GLOBALCONSTANTS OpcUaLokal (* OPC-UA-IDs fuer die lokalen Uebungen (ein Geraet) *)
  (* Standard: 61499-1; Description: Copyright (c) 2026 Meisterschulen am Ostbahnhof This program and the accompanying materials are made available under the terms of the Eclipse Public License 2.0 which is available at https://www.eclipse.org/legal/epl-2.0/ SPDX-License-Identifier: EPL-2.0 *)
  (* Version 1.0, 2026-10-18, Franz Höpfinger, Meisterschulen am Ostbahnhof, Lokal: READ/WRITE/CREATE_METHOD ohne Endpunkt, CALL_METHOD per localhost *)
  PACKAGE Meins::OPC_UA_Lokal::const;
  VAR_GLOBAL CONSTANT
    LOCAL_OPC : WSTRING := "opc.tcp://localhost:4840"; (* Eigener Server (localhost), nur fuer CALL_METHOD *)
    L01_Q1_NODE : WSTRING := "/Objects/Lokal/L01/Q1,1:s=L01_Q1"; (* L01: Knoten Q1 *)
    L01_Q1_WRITE : WSTRING := MyLib_OPC::F_OPC_LOCAL("WRITE", L01_Q1_NODE); (* L01: Input_I1 schreibt lokal (PUBLISH) *)
    L01_Q1_READ : WSTRING := MyLib_OPC::F_OPC_LOCAL("READ", L01_Q1_NODE); (* L01: Output_Q1 liest lokal (SUBSCRIBE) *)
    L03_FF1_TRIGGER_NODE : WSTRING := "/Objects/Lokal/L03/FF1_Trigger"; (* L03: Methode Toggle-Trigger *)
    L03_FF1_TRIGGER_METHOD : WSTRING := MyLib_OPC::F_OPC_LOCAL("CREATE_METHOD", L03_FF1_TRIGGER_NODE); (* L03: Methode lokal anlegen (SERVER_0) *)
    L03_FF1_TRIGGER_CALL : WSTRING := MyLib_OPC::F_OPC_REMOTE("CALL_METHOD", LOCAL_OPC, L03_FF1_TRIGGER_NODE); (* L03: Methode per localhost aufrufen (CLIENT_0) *)
    L03_FF1_STATE_NODE : WSTRING := "/Objects/Lokal/L03/FF1_State,1:s=L03_FF1_State"; (* L03: Knoten Flipflop-Zustand *)
    L03_FF1_STATE_WRITE : WSTRING := MyLib_OPC::F_OPC_LOCAL("WRITE", L03_FF1_STATE_NODE); (* L03: Zustand lokal schreiben (PUBLISH) *)
    L03_FF1_STATE_READ : WSTRING := MyLib_OPC::F_OPC_LOCAL("READ", L03_FF1_STATE_NODE); (* L03: Zustand lokal lesen (SUBSCRIBE) *)
    Q1_NODE : WSTRING := "/Objects/DigitalOutput/Q1,1:s=Output_Q1"; (* Knoten Output_Q1 *)
    Q1_READ : WSTRING := MyLib_OPC::F_OPC_LOCAL("READ", Q1_NODE); (* Output_Q1: lokal lesen (SUBSCRIBE) *)
    Q1_WRITE : WSTRING := MyLib_OPC::F_OPC_LOCAL("WRITE", Q1_NODE); (* Output_Q1: lokal schreiben (PUBLISH) *)
    FF1_TRIGGER_NODE : WSTRING := "/Objects/ToggleFF/FF1_Trigger"; (* Knoten Toggle-Trigger *)
    FF1_TRIGGER_METHOD : WSTRING := MyLib_OPC::F_OPC_LOCAL("CREATE_METHOD", FF1_TRIGGER_NODE); (* Toggle-Trigger: Methode lokal anlegen (SERVER) *)
    FF1_TRIGGER_CALL : WSTRING := MyLib_OPC::F_OPC_REMOTE("CALL_METHOD", LOCAL_OPC, FF1_TRIGGER_NODE); (* Toggle-Trigger: Methode per localhost aufrufen *)
    FF1_STATE_NODE : WSTRING := "/Objects/ToggleFF/FF1_State,1:s=FF1_State"; (* Knoten Toggle-Zustand *)
    FF1_STATE_READ : WSTRING := MyLib_OPC::F_OPC_LOCAL("READ", FF1_STATE_NODE); (* Toggle-Zustand: lokal lesen (SUBSCRIBE) *)
    FF1_STATE_WRITE : WSTRING := MyLib_OPC::F_OPC_LOCAL("WRITE", FF1_STATE_NODE); (* Toggle-Zustand: lokal schreiben (PUBLISH) *)
    SR1_SET_NODE : WSTRING := "/Objects/SRFlipflop/SR1_Set"; (* Knoten SR1 Set *)
    SR1_SET_METHOD : WSTRING := MyLib_OPC::F_OPC_LOCAL("CREATE_METHOD", SR1_SET_NODE); (* SR1 Set: Methode lokal anlegen (SERVER) *)
    SR1_SET_CALL : WSTRING := MyLib_OPC::F_OPC_REMOTE("CALL_METHOD", LOCAL_OPC, SR1_SET_NODE); (* SR1 Set: Methode per localhost aufrufen *)
    SR1_RESET_NODE : WSTRING := "/Objects/SRFlipflop/SR1_Reset"; (* Knoten SR1 Reset *)
    SR1_RESET_METHOD : WSTRING := MyLib_OPC::F_OPC_LOCAL("CREATE_METHOD", SR1_RESET_NODE); (* SR1 Reset: Methode lokal anlegen (SERVER) *)
    SR1_RESET_CALL : WSTRING := MyLib_OPC::F_OPC_REMOTE("CALL_METHOD", LOCAL_OPC, SR1_RESET_NODE); (* SR1 Reset: Methode per localhost aufrufen *)
    SR1_TOGGLE_NODE : WSTRING := "/Objects/SRFlipflop/SR1_Toggle"; (* Knoten SR1 Toggle *)
    SR1_TOGGLE_METHOD : WSTRING := MyLib_OPC::F_OPC_LOCAL("CREATE_METHOD", SR1_TOGGLE_NODE); (* SR1 Toggle: Methode lokal anlegen (SERVER) *)
    SR1_TOGGLE_CALL : WSTRING := MyLib_OPC::F_OPC_REMOTE("CALL_METHOD", LOCAL_OPC, SR1_TOGGLE_NODE); (* SR1 Toggle: Methode per localhost aufrufen *)
    SR1_STATE_NODE : WSTRING := "/Objects/SRFlipflop/SR1_State,1:s=SR1_State"; (* Knoten SR1 Zustand *)
    SR1_STATE_READ : WSTRING := MyLib_OPC::F_OPC_LOCAL("READ", SR1_STATE_NODE); (* SR1 Zustand: lokal lesen (SUBSCRIBE) *)
    SR1_STATE_WRITE : WSTRING := MyLib_OPC::F_OPC_LOCAL("WRITE", SR1_STATE_NODE); (* SR1 Zustand: lokal schreiben (PUBLISH) *)
    SR2_SET_NODE : WSTRING := "/Objects/SRFlipflop/SR2_Set"; (* Knoten SR2 Set *)
    SR2_SET_METHOD : WSTRING := MyLib_OPC::F_OPC_LOCAL("CREATE_METHOD", SR2_SET_NODE); (* SR2 Set: Methode lokal anlegen (SERVER) *)
    SR2_SET_CALL : WSTRING := MyLib_OPC::F_OPC_REMOTE("CALL_METHOD", LOCAL_OPC, SR2_SET_NODE); (* SR2 Set: Methode per localhost aufrufen *)
    SR2_RESET_NODE : WSTRING := "/Objects/SRFlipflop/SR2_Reset"; (* Knoten SR2 Reset *)
    SR2_RESET_METHOD : WSTRING := MyLib_OPC::F_OPC_LOCAL("CREATE_METHOD", SR2_RESET_NODE); (* SR2 Reset: Methode lokal anlegen (SERVER) *)
    SR2_RESET_CALL : WSTRING := MyLib_OPC::F_OPC_REMOTE("CALL_METHOD", LOCAL_OPC, SR2_RESET_NODE); (* SR2 Reset: Methode per localhost aufrufen *)
    SR2_STATE_NODE : WSTRING := "/Objects/SRFlipflop/SR2_State,1:s=SR2_State"; (* Knoten SR2 Zustand *)
    SR2_STATE_READ : WSTRING := MyLib_OPC::F_OPC_LOCAL("READ", SR2_STATE_NODE); (* SR2 Zustand: lokal lesen (SUBSCRIBE) *)
    SR2_STATE_WRITE : WSTRING := MyLib_OPC::F_OPC_LOCAL("WRITE", SR2_STATE_NODE); (* SR2 Zustand: lokal schreiben (PUBLISH) *)
    SW1_UP_NODE : WSTRING := "/Objects/Switch1/Up,1:s=Switch1_Up"; (* Knoten SW1 Hoch-Taster *)
    SW1_UP_READ : WSTRING := MyLib_OPC::F_OPC_LOCAL("READ", SW1_UP_NODE); (* SW1 Hoch-Taster: lokal lesen (SUBSCRIBE) *)
    SW1_UP_WRITE : WSTRING := MyLib_OPC::F_OPC_LOCAL("WRITE", SW1_UP_NODE); (* SW1 Hoch-Taster: lokal schreiben (PUBLISH) *)
    SW1_DOWN_NODE : WSTRING := "/Objects/Switch1/Down,1:s=Switch1_Down"; (* Knoten SW1 Runter-Taster *)
    SW1_DOWN_READ : WSTRING := MyLib_OPC::F_OPC_LOCAL("READ", SW1_DOWN_NODE); (* SW1 Runter-Taster: lokal lesen (SUBSCRIBE) *)
    SW1_DOWN_WRITE : WSTRING := MyLib_OPC::F_OPC_LOCAL("WRITE", SW1_DOWN_NODE); (* SW1 Runter-Taster: lokal schreiben (PUBLISH) *)
    SW1_UP_STATE_NODE : WSTRING := "/Objects/Switch1/UpState,1:s=Switch1_UpState"; (* Knoten SW1 Hoch erreicht *)
    SW1_UP_STATE_READ : WSTRING := MyLib_OPC::F_OPC_LOCAL("READ", SW1_UP_STATE_NODE); (* SW1 Hoch erreicht: lokal lesen (SUBSCRIBE) *)
    SW1_UP_STATE_WRITE : WSTRING := MyLib_OPC::F_OPC_LOCAL("WRITE", SW1_UP_STATE_NODE); (* SW1 Hoch erreicht: lokal schreiben (PUBLISH) *)
    SW1_DOWN_STATE_NODE : WSTRING := "/Objects/Switch1/DownState,1:s=Switch1_DownState"; (* Knoten SW1 Runter erreicht *)
    SW1_DOWN_STATE_READ : WSTRING := MyLib_OPC::F_OPC_LOCAL("READ", SW1_DOWN_STATE_NODE); (* SW1 Runter erreicht: lokal lesen (SUBSCRIBE) *)
    SW1_DOWN_STATE_WRITE : WSTRING := MyLib_OPC::F_OPC_LOCAL("WRITE", SW1_DOWN_STATE_NODE); (* SW1 Runter erreicht: lokal schreiben (PUBLISH) *)
    SW2_PRESS_NODE : WSTRING := "/Objects/Switch2/Up,1:s=Switch2_Up;/Objects/Switch2/Down,1:s=Switch2_Down"; (* Knoten SW2 Taster (2 Knoten) *)
    SW2_PRESS_READ : WSTRING := MyLib_OPC::F_OPC_LOCAL("READ", SW2_PRESS_NODE); (* SW2 Taster (2 Knoten): lokal lesen (SUBSCRIBE) *)
    SW2_PRESS_WRITE : WSTRING := MyLib_OPC::F_OPC_LOCAL("WRITE", SW2_PRESS_NODE); (* SW2 Taster (2 Knoten): lokal schreiben (PUBLISH) *)
    SW2_STATE_NODE : WSTRING := "/Objects/Switch2/UpState,1:s=Switch2_UpState;/Objects/Switch2/DownState,1:s=Switch2_DownState"; (* Knoten SW2 erreicht (2 Knoten) *)
    SW2_STATE_READ : WSTRING := MyLib_OPC::F_OPC_LOCAL("READ", SW2_STATE_NODE); (* SW2 erreicht (2 Knoten): lokal lesen (SUBSCRIBE) *)
    SW2_STATE_WRITE : WSTRING := MyLib_OPC::F_OPC_LOCAL("WRITE", SW2_STATE_NODE); (* SW2 erreicht (2 Knoten): lokal schreiben (PUBLISH) *)
    L19_Q_NODE : WSTRING := "/Objects/Lokal/L19/Q,1:s=L19_Q"; (* L19: Knoten *)
    L19_Q_WRITE : WSTRING := MyLib_OPC::F_OPC_LOCAL("WRITE", L19_Q_NODE); (* L19: Input_I1 schreibt lokal (PUBLISH) *)
    L19_Q_READ : WSTRING := MyLib_OPC::F_OPC_LOCAL("READ", L19_Q_NODE); (* L19: Output_Q1 und Output_Q2 lesen beide *)
    L13_FLIP_NODE : WSTRING := "/Objects/Lokal/L13/Flip,1:s=L13_Flip"; (* L13: Knoten Flip *)
    L13_FLOP_NODE : WSTRING := "/Objects/Lokal/L13/Flop,1:s=L13_Flop"; (* L13: Knoten Flop *)
    L13_FLIP_READ : WSTRING := MyLib_OPC::F_OPC_LOCAL("READ", L13_FLIP_NODE); (* L13: Flip lokal lesen (SUBSCRIBE) *)
    L13_FLOP_WRITE : WSTRING := MyLib_OPC::F_OPC_LOCAL("WRITE", L13_FLOP_NODE); (* L13: Flop lokal schreiben (PUBLISH) *)
    L13_FLIP_WRITE : WSTRING := MyLib_OPC::F_OPC_LOCAL("WRITE", L13_FLIP_NODE); (* L13: Input_I1 schreibt Flip lokal *)
    L13_FLOP_READ : WSTRING := MyLib_OPC::F_OPC_LOCAL("READ", L13_FLOP_NODE); (* L13: Output_Q1 liest Flop lokal *)
    L14_NUM1_NODE : WSTRING := "/Objects/Lokal/L14/Num1,1:s=L14_Num1"; (* L14: Knoten Num1 *)
    L14_NUM2_NODE : WSTRING := "/Objects/Lokal/L14/Num2,1:s=L14_Num2"; (* L14: Knoten Num2 *)
    L14_RESULT_NODE : WSTRING := "/Objects/Lokal/L14/Result,1:s=L14_Result"; (* L14: Knoten Result *)
    L14_NUM1_READ : WSTRING := MyLib_OPC::F_OPC_LOCAL("READ", L14_NUM1_NODE); (* L14: Num1 lokal lesen *)
    L14_NUM2_READ : WSTRING := MyLib_OPC::F_OPC_LOCAL("READ", L14_NUM2_NODE); (* L14: Num2 lokal lesen *)
    L14_RESULT_WRITE : WSTRING := MyLib_OPC::F_OPC_LOCAL("WRITE", L14_RESULT_NODE); (* L14: Result lokal schreiben *)
    L15_ADD_NODE : WSTRING := "/Objects/Lokal/L15/AddValues"; (* L15: Knoten AddValues *)
    L15_ADD_METHOD : WSTRING := MyLib_OPC::F_OPC_LOCAL("CREATE_METHOD", L15_ADD_NODE); (* L15: Methode AddValues anlegen (SERVER_1_2) *)
    L15_ADD_CALL : WSTRING := MyLib_OPC::F_OPC_REMOTE("CALL_METHOD", LOCAL_OPC, L15_ADD_NODE); (* L15: AddValues aufrufen (CLIENT_2_1) *)
    L16_INC_NODE : WSTRING := "/Objects/Lokal/L16/Increment,1:s=L16_Increment"; (* L16: Knoten Increment *)
    L16_INCD_NODE : WSTRING := "/Objects/Lokal/L16/Incremented,1:s=L16_Incremented"; (* L16: Knoten Incremented *)
    L16_INC_READ : WSTRING := MyLib_OPC::F_OPC_LOCAL("READ", L16_INC_NODE); (* L16: Increment lokal lesen *)
    L16_INCD_WRITE : WSTRING := MyLib_OPC::F_OPC_LOCAL("WRITE", L16_INCD_NODE); (* L16: Incremented lokal schreiben *)
    L16_INC_CLIENT_WRITE : WSTRING := MyLib_OPC::F_OPC_REMOTE("WRITE", LOCAL_OPC, L16_INC_NODE); (* L16: Increment per CLIENT schreiben *)
    L16_INCD_CLIENT_READ : WSTRING := MyLib_OPC::F_OPC_REMOTE("READ", LOCAL_OPC, L16_INCD_NODE); (* L16: Incremented per CLIENT lesen *)
    L16B_INC_NODE : WSTRING := "/Objects/Lokal/L16B/Increment,1:s=L16B_Increment"; (* L16B: Knoten Increment *)
    L16B_INCD_NODE : WSTRING := "/Objects/Lokal/L16B/Incremented,1:s=L16B_Incremented"; (* L16B: Knoten Incremented *)
    L16B_INC_READ : WSTRING := MyLib_OPC::F_OPC_LOCAL("READ", L16B_INC_NODE); (* L16B: Increment lokal lesen *)
    L16B_INCD_WRITE : WSTRING := MyLib_OPC::F_OPC_LOCAL("WRITE", L16B_INCD_NODE); (* L16B: Incremented lokal schreiben *)
    L16B_INC_CLIENT_WRITE : WSTRING := MyLib_OPC::F_OPC_REMOTE("WRITE", LOCAL_OPC, L16B_INC_NODE); (* L16B: Increment per CLIENT schreiben *)
    L16B_INCD_CLIENT_READ : WSTRING := MyLib_OPC::F_OPC_REMOTE("READ", LOCAL_OPC, L16B_INCD_NODE); (* L16B: Incremented per CLIENT lesen *)
    L17_INC_NODE : WSTRING := "/Objects/Lokal/L17/Increment,1:s=L17_Increment"; (* L17: Knoten Increment *)
    L17_INCD_NODE : WSTRING := "/Objects/Lokal/L17/Incremented,1:s=L17_Incremented"; (* L17: Knoten Incremented *)
    L17_INC_READ : WSTRING := MyLib_OPC::F_OPC_LOCAL("READ", L17_INC_NODE); (* L17: Increment lokal lesen *)
    L17_INCD_WRITE : WSTRING := MyLib_OPC::F_OPC_LOCAL("WRITE", L17_INCD_NODE); (* L17: Incremented lokal schreiben *)
    L17_INC_CLIENT_WRITE : WSTRING := MyLib_OPC::F_OPC_REMOTE("WRITE", LOCAL_OPC, L17_INC_NODE); (* L17: Increment per CLIENT schreiben *)
    L17_INCD_CLIENT_READ : WSTRING := MyLib_OPC::F_OPC_REMOTE("READ", LOCAL_OPC, L17_INCD_NODE); (* L17: Incremented per CLIENT lesen *)
    L17_INCD_SUBSCRIBE : WSTRING := MyLib_OPC::F_OPC_REMOTE("SUBSCRIBE", LOCAL_OPC, L17_INCD_NODE); (* L17: Incremented abonnieren (SUBSCRIBE mit Endpunkt) *)
    L18_OBJ_CREATE : WSTRING := "opc_ua[CREATE_OBJECT;,i=58;/Objects/1:L18_MyObject]"; (* L18: Objekt anlegen (Typ BaseObjectType i=58) *)
    L18_VAR_CREATE : WSTRING := "opc_ua[CREATE_VARIABLE;,i=63;,i=6;/Objects/1:L18_MyVariable]"; (* L18: Variable anlegen (BaseDataVariableType, Int32) *)
    L18_VAR_DELETE : WSTRING := "opc_ua[DELETE_VARIABLE;/Objects/1:L18_MyVariable]"; (* L18: Variable loeschen *)
    L18_OBJ_DELETE : WSTRING := "opc_ua[DELETE_OBJECT;/Objects/1:L18_MyObject]"; (* L18: Objekt loeschen *)
  END_VAR
END_GLOBALCONSTANTS
